Staubli VAL3: insertFOR.pgx

public program insertFOR(string x_sKey, num x_nIndex, string x_sTRAJname, num x_nLoop, string x_sIOindex, bool x_bToSave, num x_nType)
  local num l_nIndex
  local num l_i
begin

  if x_nIndex==0 and progTemp:pProgItem[x_sKey].pProgTemplate[x_nIndex].sTRAJname==""
    progTemp:pProgItem[x_sKey].pProgTemplate[x_nIndex].nType=8
    if x_nType==1
      progTemp:pProgItem[x_sKey].pProgTemplate[x_nIndex].sTRAJname="PROG"
    elseIf x_nType==2
      progTemp:pProgItem[x_sKey].pProgTemplate[x_nIndex].sTRAJname="TRAJ"
    endIf
    progTemp:pProgItem[x_sKey].pProgTemplate[x_nIndex].fForItem.sForTRAJ=x_sTRAJname
    progTemp:pProgItem[x_sKey].pProgTemplate[x_nIndex].fForItem.nLoopValue=x_nLoop
    progTemp:pProgItem[x_sKey].pProgTemplate[x_nIndex].fForItem.sIOindex=x_sIOindex
  else
    //insert(progTemp:pProgItem[x_sKey].pProgTemplate[x_nIndex+1])
    l_nIndex=x_nIndex+1
    //insert(progTemp:pProgItem[x_sKey].pProgTemplate[x_nIndex+1])
    append(progTemp:pProgItem[x_sKey].pProgTemplate)
    for l_i = size(progTemp:pProgItem[x_sKey].pProgTemplate)-1 to l_nIndex step -1
      call copyPara(x_sKey,l_i-1,l_i)
    endFor
    progTemp:pProgItem[x_sKey].pProgTemplate[x_nIndex+1].nType=8
    if x_nType==1
      progTemp:pProgItem[x_sKey].pProgTemplate[x_nIndex+1].sTRAJname="PROG"
    elseIf x_nType==2
      progTemp:pProgItem[x_sKey].pProgTemplate[x_nIndex+1].sTRAJname="TRAJ"
    endIf
    progTemp:pProgItem[x_sKey].pProgTemplate[x_nIndex+1].fForItem.sForTRAJ=x_sTRAJname
    progTemp:pProgItem[x_sKey].pProgTemplate[x_nIndex+1].fForItem.nLoopValue=x_nLoop
    progTemp:pProgItem[x_sKey].pProgTemplate[x_nIndex+1].fForItem.sIOindex=x_sIOindex
  endIf

  x_bToSave=true
end
